FUNCTION_BLOCK Gradeamento_Inovaisa (* Gradeamento mecanizado (area 100) - painel Vibropac, grades, rosca e comportas - HidrycoLib *)
  (* Standard: 61499-2 *)
  (* Version 1.1, 22/10/2026, Hidryco, Hidryco, 1.1: carga no gerador: REQ_GERADOR (geradorHabilita, stsGerador; Subestacao HAB_GM_100_01 e stsPlantaNoGerador) bloqueia o ciclo remoto na Logica e anima o raio do simbolo (AnimGerador -> STS_ANIMACAO_GERADOR). 1.0: gradeamento mecanizado da area 100 (painel Vibropac PV-35524, CLP TM241, tabela Modbus TCP Inovaisa Rev.B). Instancia "Gradeamento" com os caminhos do legado: Grade_Status1 (Controle_Gradeamento), GM_100_01/02 (Grade_Inovaisa: SensorMontante, SensorJusante, SensorDiferencial, Grade_Mecanizada_Inovaisa1), RT_100_01 (Motor_Inovaisa, rosca), CO_100_01..04 (Valvula_Coester on/off, comandadas pela IHM). Campo por symlink ${PATH}: leitura mbR4005..mbR4018 (INT), mbConexao (connStatusInt); escrita mbW4001 (ciclo), mbW4002 (reset), mbW4003/mbW4004 (setpoints 0-1000). O reset (cmdResetFalhas no E_RESET_FALHAS_PROCESSO) inclui o 4002 do painel, as grades, os sensores e as comportas. *)
  PACKAGE Hidryco.HidrycoLib;
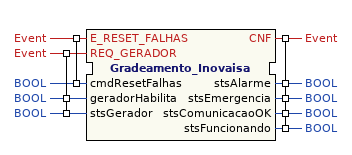
  EVENT_INPUT
    E_RESET_FALHAS WITH cmdResetFalhas; (* Reset pelo processo (painel, grades, sensores e comportas) com cmdResetFalhas = TRUE *)
    REQ_GERADOR WITH geradorHabilita, stsGerador; (* Planta no gerador e liberacao da grade (Subestacao) *)
  END_EVENT
  EVENT_OUTPUT
    CNF WITH stsAlarme, stsEmergencia, stsComunicacaoOK, stsFuncionando; (* Status *)
  END_EVENT
  VAR_INPUT
    cmdResetFalhas : BOOL; (* TRUE = reset (com o evento E_RESET_FALHAS) *)
    geradorHabilita : BOOL; (* 100-GM-01 liberada para operar com a planta nos geradores *)
    stsGerador : BOOL; (* TRUE = planta alimentada pelos geradores *)
  END_VAR
  VAR_OUTPUT
    stsAlarme : BOOL; (* Algum alarme do gradeamento (comunicacao, painel, emergencia, motores) *)
    stsEmergencia : BOOL; (* Botao de emergencia do painel acionado (4006) *)
    stsComunicacaoOK : BOOL; (* Comunicacao Modbus com o CLP do painel OK *)
    stsFuncionando : BOOL; (* Alguma grade ou a rosca funcionando *)
  END_VAR
  FBS
    IThis : Gradeamento_Inovaisa_HMI(QI := TRUE);
    plcStart1 : plcStart(Prio := 10);
    Leitura : SYMLINKMULTIVARDST_182274139AA51730B(QI := TRUE, NAME1 := '$${PATH}mbR4005', NAME2 := '$${PATH}mbR4006', NAME3 := '$${PATH}mbR4007', NAME4 := '$${PATH}mbR4008', NAME5 := '$${PATH}mbR4009', NAME6 := '$${PATH}mbR4010', NAME7 := '$${PATH}mbR4011', NAME8 := '$${PATH}mbR4012', NAME9 := '$${PATH}mbR4013', NAME10 := '$${PATH}mbR4014', NAME11 := '$${PATH}mbR4015', NAME12 := '$${PATH}mbR4016'); {SET_ATTRIBUTE(Configuration.GenericFBType.InterfaceParams, Runtime.System#I:=12;VALUE${I$}:INT,INT,INT,INT,INT,INT,INT,INT,INT,INT,INT,INT)}
    Leitura2 : SYMLINKMULTIVARDST_184BA62D721027C6E(QI := TRUE, NAME1 := '$${PATH}mbR4017', NAME2 := '$${PATH}mbR4018'); {SET_ATTRIBUTE(Configuration.GenericFBType.InterfaceParams, Runtime.System#I:=2;VALUE${I$}:INT,INT)}
    Conexao : SYMLINKMULTIVARDST_5A03F112CD5D470(QI := TRUE, NAME1 := '$${PATH}mbConexao'); {SET_ATTRIBUTE(Configuration.GenericFBType.InterfaceParams, Runtime.System#I:=1;VALUE${I$}:INT)}
    EscritaCmd : SYMLINKMULTIVARSRC_154988C56DC16E7CE(QI := TRUE, NAME1 := '$${PATH}mbW4001', NAME2 := '$${PATH}mbW4003', NAME3 := '$${PATH}mbW4004'); {SET_ATTRIBUTE(Configuration.GenericFBType.InterfaceParams, Runtime.System#I:=3;VALUE${I$}:INT,INT,INT)}
    EscritaReset : SYMLINKMULTIVARSRC_5A03F112CD5D470(QI := TRUE, NAME1 := '$${PATH}mbW4002'); {SET_ATTRIBUTE(Configuration.GenericFBType.InterfaceParams, Runtime.System#I:=1;VALUE${I$}:INT)}
    Logica : basicGradeamento;
    Tick : E_CYCLE(DT := T#1s);
    Grade_Status1 : Controle_Gradeamento;
    GM_100_01 : Grade_Inovaisa;
    GM_100_02 : Grade_Inovaisa;
    RT_100_01 : Motor_Inovaisa;
    CO_100_01 : Atuador_Coester;
    CO_100_02 : Atuador_Coester;
    CO_100_03 : Atuador_Coester;
    CO_100_04 : Atuador_Coester;
    AlarmeComunicacao : ALARM_BIT(TYPE := 1, ACKTYPE_1 := 2, ACTIVE := TRUE); {SET_ATTRIBUTE(HMI.AlarmText, Painel do gradeamento sem comunicação)} {SET_ATTRIBUTE(HMI.AlarmClass, Warning)}
    AlarmeEmergencia : ALARM_BIT(TYPE := 1, ACKTYPE_1 := 2, ACTIVE := TRUE); {SET_ATTRIBUTE(HMI.AlarmText, Emergência acionada no painel do gradeamento)}
    AlarmePainel : ALARM_BIT(TYPE := 1, ACKTYPE_1 := 2, ACTIVE := TRUE); {SET_ATTRIBUTE(HMI.AlarmText, Alarme no painel do gradeamento)}
    AnimGerador : basicCargaGerador(pin_AB02A6BAE011AA16 := TRUE);
  END_FBS
  EVENT_CONNECTIONS
    plcStart1.FIRST_INIT TO IThis.ECC090163CC0B000;
    plcStart1.REDO_INIT TO IThis.ECC090163CC0B000;
    IThis.CB22FE61A9101ECA TO Leitura.INIT;
    Leitura.INITO TO Leitura2.INIT;
    Leitura2.INITO TO Conexao.INIT;
    Conexao.INITO TO EscritaCmd.INIT;
    EscritaCmd.INITO TO EscritaReset.INIT;
    EscritaReset.INITO TO Logica.518C29172BF7055D;
    Logica.AF9623B10148EEA6 TO Tick.START;
    Leitura.CNF TO Logica.66D3215C55F0091A;
    Leitura2.CNF TO Logica.4AA0F6BC0C9CCC31;
    Conexao.CNF TO Logica.531A7DC3C1F1E4B4;
    Tick.EO TO Logica.220EF84FD56D066A;
    Grade_Status1.D0FBBC66A6D482D4 TO Logica.EAFDC5E392D9FEFA;
    Logica.9E246ABECE1E2CE6 TO Grade_Status1.BBE1950646B5A750;
    Logica.1476EEC75191AAEB TO EscritaCmd.REQ;
    Logica.1476EEC75191AAEB TO EscritaReset.REQ;
    Logica.5DAEBC207EFA920B TO GM_100_01.ABEE1148E34D9BFE;
    GM_100_01.E31D8EEC4AA83653 TO Logica.C20C38F487867904;
    Logica.5DAEBC207EFA920B TO GM_100_02.ABEE1148E34D9BFE;
    GM_100_02.E31D8EEC4AA83653 TO Logica.C20C38F487867904;
    Logica.5DAEBC207EFA920B TO RT_100_01.94DE44B005A7078D;
    RT_100_01.B512B9549703084F TO Logica.C20C38F487867904;
    IThis.242F922354BD23C9 TO Logica.6DD1F366F87AD18C;
    E_RESET_FALHAS TO Logica.D301A4C9803F7EC8;
    IThis.242F922354BD23C9 TO GM_100_01.546B340D62024106;
    IThis.242F922354BD23C9 TO GM_100_02.546B340D62024106;
    IThis.242F922354BD23C9 TO RT_100_01.86B7A273610FFA5D;
    IThis.242F922354BD23C9 TO CO_100_01.D903CD18EBE204D1;
    IThis.242F922354BD23C9 TO CO_100_02.D903CD18EBE204D1;
    IThis.242F922354BD23C9 TO CO_100_03.D903CD18EBE204D1;
    IThis.242F922354BD23C9 TO CO_100_04.D903CD18EBE204D1;
    Logica.A571F479BE4CD639 TO CNF;
    Logica.229705CA5D539927 TO IThis.38275147D3F77B46;
    Logica.229705CA5D539927 TO AlarmeComunicacao.REQ;
    AlarmeComunicacao.IND_1 TO IThis.38275147D3F77B46;
    IThis.242F922354BD23C9 TO AlarmeComunicacao.ACK_C1;
    E_RESET_FALHAS TO AlarmeComunicacao.ACK_C1;
    Logica.229705CA5D539927 TO AlarmeEmergencia.REQ;
    AlarmeEmergencia.IND_1 TO IThis.38275147D3F77B46;
    IThis.242F922354BD23C9 TO AlarmeEmergencia.ACK_C1;
    E_RESET_FALHAS TO AlarmeEmergencia.ACK_C1;
    Logica.229705CA5D539927 TO AlarmePainel.REQ;
    AlarmePainel.IND_1 TO IThis.38275147D3F77B46;
    IThis.242F922354BD23C9 TO AlarmePainel.ACK_C1;
    E_RESET_FALHAS TO AlarmePainel.ACK_C1;
    Logica.AF9623B10148EEA6 TO AlarmeComunicacao.INIT;
    AlarmeComunicacao.INITO TO AlarmeComunicacao.REQ_INITDATA;
    AlarmeComunicacao.CNF_INITDATA TO AlarmeComunicacao.ACTIVATE;
    AlarmeEmergencia.INITO TO AlarmeEmergencia.REQ_INITDATA;
    AlarmeEmergencia.CNF_INITDATA TO AlarmeEmergencia.ACTIVATE;
    AlarmeComunicacao.INITO TO AlarmeEmergencia.INIT;
    AlarmePainel.INITO TO AlarmePainel.REQ_INITDATA;
    AlarmePainel.CNF_INITDATA TO AlarmePainel.ACTIVATE;
    AlarmeEmergencia.INITO TO AlarmePainel.INIT;
    AlarmePainel.INITO TO Grade_Status1.508124526D7AA457;
    AlarmePainel.INITO TO plcStart1.ACK_FIRST;
    REQ_GERADOR TO Logica.F3638F475B575790;
    REQ_GERADOR TO AnimGerador.00789A423C908128;
    Logica.229705CA5D539927 TO AnimGerador.00789A423C908128;
    AnimGerador.D13B80EB42E4132B TO IThis.38275147D3F77B46;
  END_CONNECTIONS
  DATA_CONNECTIONS
    Leitura.VALUE1 TO Logica.EAAE7720A229695F;
    Leitura.VALUE2 TO Logica.904A23DAF55DAC59;
    Leitura.VALUE3 TO Logica.BBA94A1169D8FA73;
    Leitura.VALUE4 TO Logica.7825C7CE552E6651;
    Leitura.VALUE5 TO Logica.2498E9974464BCE6;
    Leitura.VALUE6 TO Logica.9C99F76E861BCD25;
    Leitura.VALUE7 TO Logica.D43EE0186A628319;
    Leitura.VALUE8 TO Logica.C5372D9F9D054E62;
    Leitura.VALUE9 TO Logica.9932DF3BDCD27116;
    Leitura.VALUE10 TO Logica.32562EFF83F2DC8C;
    Leitura.VALUE11 TO Logica.7C362804A2CEA9B4;
    Leitura.VALUE12 TO Logica.81F03E4BE33E3775;
    Leitura2.VALUE1 TO Logica.E74155D0A040D43B;
    Leitura2.VALUE2 TO Logica.EFE29EA2A963985E;
    Conexao.VALUE1 TO Logica.188BF646E72EEEA1;
    Grade_Status1.5789487A2939E166 TO Logica.05EA1552B9E3115E;
    Grade_Status1.8424D01B7357CBD5 TO Logica.8B073DFA930CDFDF;
    Grade_Status1.CB4F5A4E2AB68CC0 TO Logica.2CD93C02AEE34611;
    Logica.3A8B059C9015BAAF TO Grade_Status1.6CEB761D53844355;
    Logica.E8BA6941E1D9185F TO Grade_Status1.09D3C19DE8A6CC53;
    Logica.2350FEDB0EF73756 TO EscritaCmd.VALUE1;
    Logica.5A95BB21F1406E13 TO EscritaCmd.VALUE2;
    Logica.02D3ACE173D5282E TO EscritaCmd.VALUE3;
    Logica.24CB3E5A1C683D3A TO EscritaReset.VALUE1;
    Logica.B600FA4F4CE980FC TO GM_100_01.5629422A3B5B838A;
    Logica.9E07C0CEFAB1E8CD TO GM_100_01.0A48A90C6A0D0550;
    Logica.3A8B059C9015BAAF TO GM_100_01.5F90538AE86731E7;
    Logica.B48A5B93D486ADF0 TO GM_100_01.DFE6CA66F4E123D9;
    Logica.2B178368B7F1EF8F TO GM_100_01.DFA27FFCDD03BE32;
    Logica.2EE96AEBFD31A115 TO GM_100_01.550C3011667C2FB9;
    GM_100_01.7912CE47E4646D27 TO Logica.BE2397D1A1602A70;
    GM_100_01.E2890AE591C3E435 TO Logica.710DE56279147CB9;
    Logica.02DB2097D46705DB TO GM_100_02.5629422A3B5B838A;
    Logica.3E8B3064163F5CB3 TO GM_100_02.0A48A90C6A0D0550;
    Logica.E8BA6941E1D9185F TO GM_100_02.5F90538AE86731E7;
    Logica.B48A5B93D486ADF0 TO GM_100_02.DFE6CA66F4E123D9;
    Logica.4849D539B9ECCAF9 TO GM_100_02.DFA27FFCDD03BE32;
    Logica.4A2DAB6388B872A6 TO GM_100_02.550C3011667C2FB9;
    GM_100_02.7912CE47E4646D27 TO Logica.19A0761DD0428FC1;
    GM_100_02.E2890AE591C3E435 TO Logica.910F61598CD02A9A;
    Logica.A7BB4409F896B441 TO RT_100_01.7B969788E59D2A58;
    Logica.B48A5B93D486ADF0 TO RT_100_01.BC209493FBB47803;
    RT_100_01.3E3B51589C07F168 TO Logica.A295421A8158BEBA;
    RT_100_01.9F7A867A79CFF3D0 TO Logica.373787043AB8D8D4;
    IThis.6A21846A09042795 TO Logica.C648B0BD976A65D6;
    cmdResetFalhas TO Logica.E2508CD3A47CDCD2;
    IThis.6A21846A09042795 TO GM_100_01.605D63048CED98E9;
    IThis.6A21846A09042795 TO GM_100_02.605D63048CED98E9;
    IThis.6A21846A09042795 TO RT_100_01.08D30EE79B49C6AD;
    IThis.6A21846A09042795 TO CO_100_01.C82CBBE25FC56079;
    IThis.6A21846A09042795 TO CO_100_02.C82CBBE25FC56079;
    IThis.6A21846A09042795 TO CO_100_03.C82CBBE25FC56079;
    IThis.6A21846A09042795 TO CO_100_04.C82CBBE25FC56079;
    Logica.8A40AFCE6F808DC2 TO stsAlarme;
    Logica.D4E1CE246816215C TO stsEmergencia;
    Logica.D2C98E15D329182A TO stsComunicacaoOK;
    Logica.F73DC825969A7AAC TO stsFuncionando;
    Logica.8A40AFCE6F808DC2 TO IThis.6FCA39A2D147DE77;
    Logica.D4E1CE246816215C TO IThis.F045091C645F3312;
    Logica.D2C98E15D329182A TO IThis.5A984024F490CFC5;
    Logica.B069C22B63DCD037 TO IThis.39BED905FADF3373;
    Logica.4914469ABA3CB0F5 TO IThis.A5523AEDFD3969A6;
    Logica.26FB5E58803038CB TO IThis.51D5459D1498110E;
    Logica.77ADF001A8F11DA2 TO IThis.1D655E340905F44F;
    Logica.F73DC825969A7AAC TO IThis.9512D253D4D322C2;
    Logica.B069C22B63DCD037 TO AlarmeComunicacao.INP;
    AlarmeComunicacao.STATE_1 TO IThis.4E0788183C903F3D;
    Logica.D4E1CE246816215C TO AlarmeEmergencia.INP;
    AlarmeEmergencia.STATE_1 TO IThis.27D2486D2537D0D5;
    Logica.4914469ABA3CB0F5 TO AlarmePainel.INP;
    AlarmePainel.STATE_1 TO IThis.9BCF8DFF4840D2B4;
    geradorHabilita TO Logica.162C592D6763A41A;
    stsGerador TO Logica.29083538F3254FDC;
    geradorHabilita TO AnimGerador.E98CC3FC79967C8B;
    stsGerador TO AnimGerador.9DDD74C1F0C45B78;
    Logica.F73DC825969A7AAC TO AnimGerador.92CF573A93E227B1;
    AnimGerador.87DFF1D389B6D369 TO IThis.4B4EC1B0C0F9D0FF;
  END_CONNECTIONS
END_FUNCTION_BLOCK
